(* IEC 61131-3 sources: ST-graph-rag-mcp/test/fixtures/c2-test, 1 file *)

(* ---- FB_Test.st ---- *)
FUNCTION_BLOCK FB_Test
VAR_INPUT x : BOOL; END_VAR
END_FUNCTION_BLOCK
